--- program DoorRL_C (robot ABB IRB 1300-10/1.15) ---
  Smooth(1)
  Set speed (1000.0 mm/s)
  Set Ref.: DoorRL
  Set Tool: Generic Paint Sprayer
  Show Generic Paint Sprayer
  MoveJ 1 to (90.7, 0.32, 7.32) mm, rotated rx -9.04 ry 0.01 rz 91.21 deg; joints [83.599, -28.806, 2.512, -49.508, 32.312, -224.781, 2064.306, 3452.351, 803.193]
  MoveL 2 to (90.7, 0.32, 7.32) mm, rotated rx -9.04 ry 0.01 rz 91.21 deg; joints [83.599, -28.806, 2.512, -49.508, 32.312, -224.781, 2064.306, 3452.351, 803.193]
  MoveL 3 to (75, 0, 106.08) mm, rotated rx -9.04 ry 0.01 rz 91.21 deg; joints [85.387, -19.776, -1.909, -57.854, 30.896, -215.842, 2064.306, 3452.351, 803.193]
  MoveL 4 to (75, 0, 106.08) mm, rotated rx -9.04 ry 0.01 rz 91.21 deg; joints [85.387, -19.776, -1.909, -57.854, 30.896, -215.842, 2064.306, 3452.351, 803.193]
  Set speed (200.0 mm/s)
  MoveL 5 to (75, 100, 106.62) mm, rotated rx -8.72 ry -0.14 rz 91.23 deg; joints [102.46, -18.99, -2.4, -72.728, 45.516, -205.072, 2064.306, 3452.351, 803.193]
  MoveL 6 to (75, 200, 107.42) mm, rotated rx -8.48 ry -0.48 rz 91.28 deg; joints [117.629, -15.548, -4.305, -81.612, 59.424, -199.395, 2064.306, 3452.351, 803.193]
  MoveL 7 to (75, 300, 108.62) mm, rotated rx -8.1 ry -0.62 rz 91.29 deg; joints [129.26, -10.149, -8.101, -86.402, 70.427, -196.705, 2064.306, 3452.351, 803.193]
  MoveL 8 to (75, 400, 110.17) mm, rotated rx -8.3 ry -0.88 rz 91.34 deg; joints [137.912, -3.315, -13.206, -89.791, 78.836, -194.463, 2064.306, 3452.351, 803.193]
  MoveL 9 to (75, 500, 112.34) mm, rotated rx -7.79 ry -1.35 rz 91.39 deg; joints [144.305, 5.186, -22.224, -91.259, 85.516, -195.347, 2064.306, 3452.351, 803.193]
  MoveL 10 to (75, 600, 114.4) mm, rotated rx -6.61 ry -0.07 rz 91.2 deg; joints [148.976, 13.47, -33.602, -91.242, 88.944, -199.214, 2064.306, 3452.351, 803.193]
  Set speed (1000.0 mm/s)
  MoveL 11 to (75, 600, 114.4) mm, rotated rx -6.61 ry -0.07 rz 91.2 deg; joints [148.976, 13.47, -33.602, -91.242, 88.944, -199.214, 2064.306, 3452.351, 803.193]
  MoveL 12 to (86.51, 600.37, 15.07) mm, rotated rx -6.61 ry -0.07 rz 91.2 deg; joints [156.899, 8.317, -26.551, -93.775, 96.503, -197.647, 2064.306, 3452.351, 803.193]
  Set speed (1000.0 mm/s)
  MoveL 13 to (152.01, 598.2, 20.45) mm, rotated rx -1.13 ry 1.05 rz 91.14 deg; joints [156.743, 6.079, -21.228, -88.467, 96.739, -196.702, 2064.306, 3452.351, 803.193]
  MoveL 14 to (150, 600, 120.41) mm, rotated rx -1.13 ry 1.05 rz 91.14 deg; joints [148.769, 10.819, -26.045, -86.396, 89.056, -197.123, 2064.306, 3452.351, 803.193]
  MoveL 15 to (150, 600, 120.41) mm, rotated rx -1.13 ry 1.05 rz 91.14 deg; joints [148.769, 10.819, -26.045, -86.396, 89.056, -197.123, 2064.306, 3452.351, 803.193]
  Set speed (200.0 mm/s)
  MoveL 16 to (150, 500, 121.61) mm, rotated rx -2.1 ry 0.62 rz 91.14 deg; joints [143.656, 2.312, -15.23, -86.198, 84.142, -194.609, 2064.306, 3452.351, 803.193]
  MoveL 17 to (150, 400, 121.47) mm, rotated rx -4.4 ry -0.1 rz 91.19 deg; joints [137.209, -5.289, -5.416, -87.296, 77.972, -191.254, 2064.306, 3452.351, 803.193]
  MoveL 18 to (150, 300, 120.53) mm, rotated rx -8.5 ry -0.52 rz 91.29 deg; joints [128.581, -12.398, 4.736, -90.48, 69.312, -185.121, 2064.306, 3452.351, 803.193]
  MoveL 19 to (150, 200, 119.49) mm, rotated rx -8.12 ry -0.38 rz 91.26 deg; joints [116.951, -17.771, 7.428, -86.802, 57.781, -188.768, 2064.306, 3452.351, 803.193]
  MoveL 20 to (150, 100, 118.81) mm, rotated rx -7.65 ry -0.05 rz 91.21 deg; joints [101.911, -21.13, 8.356, -79.735, 43.178, -194.732, 2064.306, 3452.351, 803.193]
  MoveL 21 to (150, 0, 118.53) mm, rotated rx -7.91 ry 0.3 rz 91.16 deg; joints [84.752, -21.907, 8.755, -69.015, 26.732, -202.933, 2064.306, 3452.351, 803.193]
  Set speed (1000.0 mm/s)
  MoveL 22 to (150, 0, 118.53) mm, rotated rx -7.91 ry 0.3 rz 91.16 deg; joints [84.752, -21.907, 8.755, -69.015, 26.732, -202.933, 2064.306, 3452.351, 803.193]
  MoveL 23 to (163.76, -0.24, 19.48) mm, rotated rx -7.91 ry 0.3 rz 91.16 deg; joints [82.61, -31.376, 12.865, -57.206, 27.32, -215.521, 2064.306, 3452.351, 803.193]
  Set speed (1000.0 mm/s)
  MoveL 24 to (223.66, 0.79, 20.64) mm, rotated rx 0.76 ry -0.47 rz 91.14 deg; joints [84.141, -30.772, 10.615, -47.345, 35.088, -229.019, 2064.306, 3452.351, 803.193]
  MoveL 25 to (225, 0, 120.63) mm, rotated rx 0.76 ry -0.47 rz 91.14 deg; joints [85.606, -21.929, 8.883, -57.612, 31.856, -217.231, 2064.306, 3452.351, 803.193]
  MoveL 26 to (225, 0, 120.63) mm, rotated rx 0.76 ry -0.47 rz 91.14 deg; joints [85.606, -21.929, 8.883, -57.612, 31.856, -217.231, 2064.306, 3452.351, 803.193]
  Set speed (200.0 mm/s)
  MoveL 27 to (225, 100, 121.28) mm, rotated rx 0.7 ry -0.35 rz 91.14 deg; joints [102.099, -21.314, 8.944, -70.725, 45.982, -205.135, 2064.306, 3452.351, 803.193]
  MoveL 28 to (225, 200, 122.15) mm, rotated rx 0.5 ry -0.52 rz 91.15 deg; joints [117.028, -17.979, 7.742, -78.485, 59.657, -197.425, 2064.306, 3452.351, 803.193]
  MoveL 29 to (225, 300, 123.05) mm, rotated rx 0.21 ry -0.42 rz 91.15 deg; joints [128.604, -12.816, 5.114, -82.577, 70.367, -192.361, 2064.306, 3452.351, 803.193]
  MoveL 30 to (225, 400, 123.5) mm, rotated rx -0.2 ry -0.26 rz 91.16 deg; joints [137.37, -6.35, 0.883, -84.796, 78.558, -188.773, 2064.306, 3452.351, 803.193]
  MoveL 31 to (225, 500, 123.04) mm, rotated rx -1.05 ry 0.5 rz 91.15 deg; joints [143.943, 0.436, -4.189, -86.301, 84.114, -186.009, 2064.306, 3452.351, 803.193]
  MoveL 32 to (225, 600, 122.08) mm, rotated rx -1.6 ry 0.73 rz 91.14 deg; joints [149.099, 8.52, -12.229, -87.11, 88.967, -185.37, 2064.306, 3452.351, 803.193]
  MoveL 33 to (225, 700, 120.88) mm, rotated rx 0.16 ry -3.32 rz 91.14 deg; joints [153.063, 22.747, -33.337, -87.148, 97.49, -192.931, 2064.306, 3452.351, 803.193]
  Set speed (1000.0 mm/s)
  MoveL 34 to (225, 700, 120.88) mm, rotated rx 0.16 ry -3.32 rz 91.14 deg; joints [153.063, 22.747, -33.337, -87.148, 97.49, -192.931, 2064.306, 3452.351, 803.193]
  MoveL 35 to (224.61, 705.78, 21.05) mm, rotated rx 0.16 ry -3.32 rz 91.14 deg; joints [160.083, 19.015, -28.957, -88.222, 104.365, -191.988, 2064.306, 3452.351, 803.193]
  Set speed (1000.0 mm/s)
  MoveL 36 to (305.54, 698.73, 24.64) mm, rotated rx -3.16 ry 0.79 rz 91.13 deg; joints [160.573, 12.44, -5.322, -87.261, 99.896, -173.342, 2064.306, 3452.351, 803.193]
  MoveL 37 to (300, 700, 124.48) mm, rotated rx -3.16 ry 0.79 rz 91.13 deg; joints [153.278, 16.534, -10.403, -88.244, 92.694, -174.618, 2064.306, 3452.351, 803.193]
  MoveL 38 to (300, 700, 124.48) mm, rotated rx -3.16 ry 0.79 rz 91.13 deg; joints [153.278, 16.534, -10.403, -88.244, 92.694, -174.618, 2064.306, 3452.351, 803.193]
  Set speed (200.0 mm/s)
  MoveL 39 to (300, 600, 125.06) mm, rotated rx -3.23 ry 0.19 rz 91.16 deg; joints [149.376, 8.214, 0.141, -88.693, 89.372, -172.462, 2064.306, 3452.351, 803.193]
  MoveL 40 to (300, 500, 125.16) mm, rotated rx -2.17 ry 0.14 rz 91.16 deg; joints [144.303, -0.143, 7.785, -88.428, 84.307, -173.89, 2064.306, 3452.351, 803.193]
  MoveL 41 to (300, 400, 124.72) mm, rotated rx -1.66 ry -0.34 rz 91.17 deg; joints [137.782, -7.551, 13.671, -88.464, 78.321, -175.937, 2064.306, 3452.351, 803.193]
  MoveL 42 to (300, 300, 123.67) mm, rotated rx -1.09 ry -0.54 rz 91.17 deg; joints [129.056, -14.44, 17.858, -87.824, 69.893, -179.463, 2064.306, 3452.351, 803.193]
  MoveL 43 to (300, 200, 122.54) mm, rotated rx -1.3 ry -0.63 rz 91.18 deg; joints [117.411, -20.166, 21.239, -87.099, 58.454, -182.429, 2064.306, 3452.351, 803.193]
  MoveL 44 to (300, 100, 121.57) mm, rotated rx -1.33 ry -0.43 rz 91.17 deg; joints [102.223, -23.973, 22.85, -84.399, 43.259, -186.653, 2064.306, 3452.351, 803.193]
  MoveL 45 to (300, 0, 120.78) mm, rotated rx -1.5 ry -0.32 rz 91.17 deg; joints [85.014, -24.825, 23.131, -79.981, 26.14, -191.455, 2064.306, 3452.351, 803.193]
  Set speed (1000.0 mm/s)
  MoveL 46 to (300, 0, 120.78) mm, rotated rx -1.5 ry -0.32 rz 91.17 deg; joints [85.014, -24.825, 23.131, -79.981, 26.14, -191.455, 2064.306, 3452.351, 803.193]
  MoveL 47 to (302.6, 0.61, 20.82) mm, rotated rx -1.5 ry -0.32 rz 91.17 deg; joints [83.173, -35.007, 25.553, -63.775, 26.819, -209.331, 2064.306, 3452.351, 803.193]
  Set speed (1000.0 mm/s)
  MoveL 48 to (382.47, 0.73, 24.79) mm, rotated rx -4.29 ry -0.33 rz 91.21 deg; joints [82.724, -37.124, 40.086, -95.64, 23.549, -173.926, 2064.306, 3452.351, 803.193]
  MoveL 49 to (375, 0, 124.51) mm, rotated rx -4.29 ry -0.33 rz 91.21 deg; joints [84.717, -25.281, 36.632, -111.575, 27.492, -156.03, 2064.306, 3452.351, 803.193]
  MoveL 50 to (375, 0, 124.51) mm, rotated rx -4.29 ry -0.33 rz 91.21 deg; joints [84.717, -25.281, 36.632, -111.575, 27.492, -156.03, 2064.306, 3452.351, 803.193]
  Set speed (200.0 mm/s)
  MoveL 51 to (375, 100, 125.3) mm, rotated rx -4.19 ry -0.39 rz 91.21 deg; joints [102.046, -24.392, 36.412, -101.899, 43.99, -163.49, 2064.306, 3452.351, 803.193]
  MoveL 52 to (375, 200, 126.3) mm, rotated rx -3.97 ry -0.6 rz 91.22 deg; joints [117.418, -20.181, 34.415, -97.776, 59.26, -164.282, 2064.306, 3452.351, 803.193]
  MoveL 53 to (375, 300, 127.56) mm, rotated rx -5.31 ry -0.62 rz 91.24 deg; joints [129.232, -13.59, 32.312, -96.985, 71.452, -159.822, 2064.306, 3452.351, 803.193]
  MoveL 54 to (375, 400, 128.83) mm, rotated rx -5.27 ry -0.59 rz 91.24 deg; joints [137.993, -6.109, 26.861, -94.307, 79.819, -158.606, 2064.306, 3452.351, 803.193]
  MoveL 55 to (375, 500, 129.91) mm, rotated rx -4.47 ry -0.21 rz 91.2 deg; joints [144.445, 1.382, 19.151, -91.452, 85.235, -159.606, 2064.306, 3452.351, 803.193]
  MoveL 56 to (375, 600, 130.48) mm, rotated rx -5.59 ry -0.1 rz 91.2 deg; joints [149.411, 9.838, 11.165, -90.644, 90.13, -158.616, 2064.306, 3452.351, 803.193]
  MoveL 57 to (375, 700, 130.64) mm, rotated rx -6.1 ry 0.33 rz 91.16 deg; joints [153.257, 18.109, 1.02, -89.952, 93.484, -160.267, 2064.306, 3452.351, 803.193]
  MoveL 58 to (375, 800, 129.84) mm, rotated rx -6.14 ry 1.82 rz 91 deg; joints [156.376, 25.705, -10.148, -89.777, 95.052, -163.863, 2064.306, 3452.351, 803.193]
  Set speed (1000.0 mm/s)
  MoveL 59 to (375, 800, 129.84) mm, rotated rx -6.14 ry 1.82 rz 91 deg; joints [156.376, 25.705, -10.148, -89.777, 95.052, -163.863, 2064.306, 3452.351, 803.193]
  MoveL 60 to (385.74, 797.03, 30.46) mm, rotated rx -6.14 ry 1.82 rz 91 deg; joints [163.022, 22.035, -4.129, -87.501, 101.36, -161.341, 2064.306, 3452.351, 803.193]
  Set speed (1000.0 mm/s)
  MoveL 61 to (473.75, 798.92, 46.41) mm, rotated rx -13.73 ry 0.89 rz 91.03 deg; joints [161.964, 28.907, 7.054, -89.444, 104.008, -140.367, 2064.306, 3452.351, 803.193]
  MoveL 62 to (450, 800, 143.54) mm, rotated rx -13.73 ry 0.89 rz 91.03 deg; joints [155.503, 31.395, 0.291, -93.866, 98.516, -144.558, 2064.306, 3452.351, 803.193]
  MoveL 63 to (450, 800, 143.54) mm, rotated rx -13.73 ry 0.89 rz 91.03 deg; joints [155.503, 31.395, 0.291, -93.866, 98.516, -144.558, 2064.306, 3452.351, 803.193]
  Set speed (200.0 mm/s)
  MoveL 64 to (450, 700, 143.19) mm, rotated rx -13.87 ry 0.24 rz 91.18 deg; joints [152.373, 24.011, 12.763, -94.602, 96.91, -139.132, 2064.306, 3452.351, 803.193]
  MoveL 65 to (450, 600, 141.71) mm, rotated rx -14.05 ry -0.52 rz 91.38 deg; joints [148.554, 17.067, 23.436, -96.144, 94.968, -134.987, 2064.306, 3452.351, 803.193]
  MoveL 66 to (450, 500, 140.16) mm, rotated rx -13.37 ry -0.76 rz 91.42 deg; joints [143.712, 9.342, 32.755, -98.644, 91.321, -133.254, 2064.306, 3452.351, 803.193]
  MoveL 67 to (450, 400, 138.58) mm, rotated rx -12.7 ry -0.52 rz 91.35 deg; joints [137.185, 1.179, 40.884, -102.834, 85.962, -132.737, 2064.306, 3452.351, 803.193]
  MoveL 68 to (450, 300, 137.1) mm, rotated rx -11.58 ry -0.68 rz 91.37 deg; joints [128.567, -6.84, 46.323, -107.585, 78.404, -134.195, 2064.306, 3452.351, 803.193]
  MoveL 69 to (450, 200, 135.73) mm, rotated rx -11.11 ry -0.72 rz 91.37 deg; joints [116.912, -13.706, 50.251, -114.63, 68.528, -133.929, 2064.306, 3452.351, 803.193]
  MoveL 70 to (450, 100, 134.52) mm, rotated rx -9.69 ry -0.28 rz 91.26 deg; joints [101.492, -19.511, 51.351, -123.947, 53.928, -132.478, 2064.306, 3452.351, 803.193]
  MoveL 71 to (450, 0, 133.84) mm, rotated rx -9.43 ry -0.15 rz 91.24 deg; joints [84.256, -20.688, 51.274, -141.098, 41.917, -120.478, 2064.306, 3452.351, 803.193]
  Set speed (1000.0 mm/s)
  MoveL 72 to (450, 0, 133.84) mm, rotated rx -9.43 ry -0.15 rz 91.24 deg; joints [84.256, -20.688, 51.274, -141.098, 41.917, -120.478, 2064.306, 3452.351, 803.193]
  MoveL 73 to (466.37, 0.62, 35.19) mm, rotated rx -9.43 ry -0.15 rz 91.24 deg; joints [82.039, -34.232, 56.958, -137.497, 34.657, -126.322, 2064.306, 3452.351, 803.193]
  Set speed (1000.0 mm/s)
  MoveL 74 to (555.05, -82.25, 116.77) mm, rotated rx 60.29 ry -13.07 rz -152.57 deg; joints [70.284, 61.29, -33.097, 77.942, 86.027, -269.551, 2564.306, 3828.918, 1060.29]
  MoveL 75 to (525, 0, 165.05) mm, rotated rx 37.44 ry 52.55 rz 154.03 deg; joints [24.866, 61.421, -22.556, 79.321, 94.582, -359.342, 1755.93, 3452.351, 1099.978]
  MoveL 76 to (525, 0, 165.05) mm, rotated rx 37.44 ry 52.55 rz 154.03 deg; joints [24.866, 61.421, -22.556, 79.321, 94.582, -359.342, 1755.93, 3452.351, 1099.978]
  Set speed (200.0 mm/s)
  MoveL 77 to (525, 100, 155.04) mm, rotated rx -9.84 ry 16.5 rz 149.85 deg; joints [40.939, 27.228, 59.96, 145.73, 75.776, -387.964, 1755.93, 3452.351, 1099.978]
  MoveL 78 to (525, 200, 156.11) mm, rotated rx 15.18 ry 12.68 rz -126.97 deg; joints [110.817, 44.311, 23.812, 178.664, 63.101, -311.328, 2564.306, 3828.918, 1099.979]
  MoveL 79 to (525, 300, 157.73) mm, rotated rx -8.79 ry -16.06 rz 32.63 deg; joints [133.225, 83.406, -21.75, 229.016, 112.204, -168.506, 2564.306, 3742.832, 1099.974]
  MoveL 80 to (525, 400, 159.79) mm, rotated rx -8.89 ry -16.44 rz 32.7 deg; joints [137.126, 86.051, -37.16, 228.381, 105.823, -180.156, 2564.306, 3742.832, 1060.252]
  MoveL 81 to (525, 500, 162.03) mm, rotated rx -9.11 ry -16.87 rz 32.78 deg; joints [140.443, 100.168, -72.983, 227.152, 93.486, -198.143, 2564.306, 3742.832, 1060.252]
  MoveL 82 to (525, 600, 164.37) mm, rotated rx -9.81 ry -18.17 rz 33.04 deg; joints [119.482, 84.102, -18.159, 219.568, 113.288, -160.148, 2064.306, 3834.482, 1099.978]
  MoveL 83 to (525, 700, 166.85) mm, rotated rx -10.72 ry -19.05 rz 33.23 deg; joints [124.134, 85.187, -28.709, 220.198, 108.523, -168.206, 2064.306, 3834.482, 1060.086]
  MoveL 84 to (525, 800, 169.19) mm, rotated rx -11.61 ry -20.92 rz 33.67 deg; joints [131.809, 86.524, -29.394, 225.322, 113.849, -170.732, 2064.306, 3735.345, 1060.086]
  MoveL 85 to (525, 900, 171.75) mm, rotated rx -12.62 ry -22.91 rz 34.2 deg; joints [135.296, 97.473, -57.469, 222.496, 105.147, -184.837, 2064.306, 3735.345, 1060.086]
  Set speed (1000.0 mm/s)
  MoveL 86 to (525, 900, 171.75) mm, rotated rx -12.62 ry -22.91 rz 34.2 deg; joints [135.296, 97.473, -57.469, 222.496, 105.147, -184.837, 2064.306, 3735.345, 1060.086]
  MoveL 87 to (568.69, 903.29, 81.86) mm, rotated rx -12.62 ry -22.91 rz 34.2 deg; joints [135.12, 104.561, -69.901, 221.579, 101.084, -188.404, 2064.306, 3836.185, 1060.086]
  Set speed (1000.0 mm/s)
  MoveL 88 to (674.57, 902.94, 144.38) mm, rotated rx -46.41 ry -15.12 rz 78.31 deg; joints [105.449, 76.927, -11.434, 224.156, 120.066, -102.909, 1454.359, 3827.063, 803.193]
  MoveL 89 to (600, 900, 210.95) mm, rotated rx -46.41 ry -15.12 rz 78.31 deg; joints [105.243, 71.137, -8.955, 222.754, 117.599, -105.433, 1454.359, 3760.201, 803.193]
  MoveL 90 to (600, 900, 210.95) mm, rotated rx -46.41 ry -15.12 rz 78.31 deg; joints [105.243, 71.137, -8.955, 222.754, 117.599, -105.433, 1454.359, 3760.201, 803.193]
  Set speed (200.0 mm/s)
  MoveL 91 to (600, 800, 210) mm, rotated rx 6.16 ry 2.87 rz 71.3 deg; joints [100.8, 46.533, 29.485, 219.508, 78.715, -121.802, 1454.359, 3760.201, 1056.724]
  MoveL 92 to (600, 700, 203.49) mm, rotated rx -43.73 ry -14.25 rz 77.35 deg; joints [92.704, 90.414, -14.669, 216.98, 122.816, -93.221, 1454.359, 3760.201, 1056.724]
  MoveL 93 to (600, 600, 200.56) mm, rotated rx -44.05 ry -14.06 rz 77.17 deg; joints [85.887, 90.364, -14.403, 211.003, 122.369, -91.43, 1454.359, 3760.201, 1056.724]
  MoveL 94 to (600, 500, 198.23) mm, rotated rx -43.4 ry -13.95 rz 77.05 deg; joints [79.336, 89.984, -14.885, 205.125, 120.303, -90.613, 1454.359, 3760.201, 1056.724]
  MoveL 95 to (600, 400, 196.18) mm, rotated rx -44.51 ry 0.19 rz 91.33 deg; joints [104.974, 82.58, -3.734, 227.238, 116.231, -77.118, 1920.961, 3772.068, 1056.724]
  MoveL 96 to (600, 300, 194.65) mm, rotated rx -43.34 ry 0.41 rz 91.12 deg; joints [98.134, 80.928, 1.713, 221.6, 117.257, -74.136, 1920.961, 3772.068, 1056.724]
  MoveL 97 to (600, 200, 193.74) mm, rotated rx -42.2 ry 0.55 rz 90.99 deg; joints [90.952, 79.687, 4.868, 214.872, 117.373, -72.904, 1920.961, 3772.068, 1056.724]
  MoveL 98 to (600, 100, 193.19) mm, rotated rx -40.28 ry 0.54 rz 91.01 deg; joints [83.708, 78.061, 6.898, 207.528, 115.777, -73.221, 1920.961, 3772.068, 1056.724]
  Set speed (1000.0 mm/s)
  MoveL 99 to (600, 100, 193.19) mm, rotated rx -40.28 ry 0.54 rz 91.01 deg; joints [83.708, 78.061, 6.898, 207.528, 115.777, -73.221, 1920.961, 3772.068, 1056.724]
  MoveL 100 to (664.66, 100.42, 116.91) mm, rotated rx -40.28 ry 0.54 rz 91.01 deg; joints [83.431, 83.386, 6.777, 208.563, 120.365, -70.437, 1920.961, 3823.518, 1056.724]
  Set speed (1000.0 mm/s)
  MoveL 101 to (748.8, 402.34, 190.34) mm, rotated rx -47.59 ry -0.13 rz 91.7 deg; joints [105.259, 99.236, -20.482, 228.709, 118.671, -75.099, 1920.961, 3768.591, 1056.724]
  MoveL 102 to (675, 400, 257.78) mm, rotated rx -47.59 ry -0.13 rz 91.7 deg; joints [103.965, 94.987, -25.674, 224.332, 111.906, -82.4, 1920.961, 3768.591, 1056.724]
  MoveL 103 to (675, 400, 257.78) mm, rotated rx -47.59 ry -0.13 rz 91.7 deg; joints [103.965, 94.987, -25.674, 224.332, 111.906, -82.4, 1920.961, 3768.591, 1056.724]
  Set speed (200.0 mm/s)
  MoveL 104 to (675, 500, 261.5) mm, rotated rx -47.59 ry -0.25 rz 91.84 deg; joints [109.884, 97.185, -33.463, 227.815, 109.711, -88.385, 1920.961, 3768.591, 1056.724]
  MoveL 105 to (675, 600, 265.72) mm, rotated rx -44.04 ry -14.72 rz 77.83 deg; joints [86.509, 101.363, -35.436, 209.841, 113.733, -96.969, 1454.359, 3755.143, 1056.724]
  MoveL 106 to (675, 700, 270.37) mm, rotated rx -41.7 ry -14.36 rz 77.4 deg; joints [92.877, 99.524, -31.623, 214.934, 114.764, -99.411, 1454.359, 3755.143, 1056.724]
  MoveL 107 to (675, 800, 275.52) mm, rotated rx -37.38 ry -13.59 rz 76.58 deg; joints [99.465, 96.499, -26.735, 220.282, 114.038, -102.592, 1454.359, 3755.143, 1056.724]
  MoveL 108 to (675, 900, 280.97) mm, rotated rx -37.72 ry -1.38 rz 92.5 deg; joints [104.161, 95.633, -32.168, 224.415, 99.282, -91.601, 1420.961, 3825.258, 1099.805]
  MoveL 109 to (675, 1000, 287.24) mm, rotated rx -31.01 ry -12.9 rz 75.77 deg; joints [112.266, 94.902, -31.121, 229.795, 108.116, -113.99, 1454.359, 3755.143, 1056.724]
  Set speed (1000.0 mm/s)
  MoveL 110 to (675, 1000, 287.24) mm, rotated rx -31.01 ry -12.9 rz 75.77 deg; joints [112.266, 94.902, -31.121, 229.795, 108.116, -113.99, 1454.359, 3755.143, 1056.724]
  MoveL 111 to (729.64, 1005.88, 203.7) mm, rotated rx -25.34 ry -22.43 rz 57.28 deg; joints [118.128, 111.273, -49.466, 227.376, 116.936, -137.304, 1564.306, 3749.389, 1099.805]

--- program DoorFL_C (robot ABB IRB 1300-10/1.15) ---
  Smooth(1)
  Set speed (1000.0 mm/s)
  Set Ref.: DoorFL
  Set Tool: Generic Paint Sprayer
  Show Generic Paint Sprayer
  MoveJ 1 to (71.29, 9.92, 20.7) mm, rotated rx 1.8 ry -5.81 rz 93.26 deg; joints [-42.65, -30.194, 5.671, 93.562, 99.411, 24.312, 2956.487, 3047.951, 891.281]
  MoveL 2 to (71.29, 9.92, 20.7) mm, rotated rx 1.8 ry -5.81 rz 93.26 deg; joints [-42.65, -30.194, 5.671, 93.562, 99.411, 24.312, 2956.487, 3047.951, 891.281]
  MoveL 3 to (75, 0, 120.14) mm, rotated rx 1.8 ry -5.81 rz 93.26 deg; joints [-42.65, -30.194, 5.671, 93.562, 99.411, 24.312, 2961.047, 2948.065, 889.846]
  MoveL 4 to (75, 0, 120.14) mm, rotated rx 1.8 ry -5.81 rz 93.26 deg; joints [-42.65, -30.194, 5.671, 93.562, 99.411, 24.312, 2961.047, 2948.065, 889.846]
  Set speed (200.0 mm/s)
  MoveL 5 to (75, 100, 126.97) mm, rotated rx -3.91 ry -2.93 rz 93.33 deg; joints [-42.529, -30.194, 9.554, 98.562, 100.324, 24.312, 2875.19, 2948.065, 860.651]
  MoveL 6 to (75, 200, 131.93) mm, rotated rx -5.64 ry -2.28 rz 93.25 deg; joints [-42.357, -30.194, 10.675, 99.97, 100.324, 24.312, 2777.783, 2947.743, 847.202]
  MoveL 7 to (75, 300, 136.32) mm, rotated rx -5.77 ry -2.17 rz 93.24 deg; joints [-42.357, -30.194, 10.767, 100.106, 100.386, 24.312, 2678.543, 2948.883, 840.768]
  MoveL 8 to (75, 400, 140.74) mm, rotated rx -5.66 ry -2.28 rz 93.25 deg; joints [-42.432, -30.263, 10.767, 100.006, 100.386, 24.312, 2578.494, 2949.946, 835.842]
  MoveL 9 to (75, 500, 145.36) mm, rotated rx -5.57 ry -2.46 rz 93.27 deg; joints [-42.582, -30.306, 10.767, 99.924, 100.386, 24.312, 2477.83, 2950.073, 830.733]
  MoveL 10 to (75, 600, 150.28) mm, rotated rx -5.46 ry -2.6 rz 93.29 deg; joints [-42.694, -30.37, 10.767, 99.824, 100.386, 24.312, 2377.497, 2950.334, 825.812]
  MoveL 11 to (75, 700, 155.46) mm, rotated rx -5.27 ry -2.81 rz 93.31 deg; joints [-42.844, -30.483, 10.767, 99.658, 100.386, 24.312, 2277.163, 2950.452, 821.515]
  MoveL 12 to (75, 800, 160.96) mm, rotated rx -5.04 ry -2.89 rz 93.32 deg; joints [-42.859, -30.634, 10.767, 99.472, 100.386, 24.312, 2177.86, 2951.505, 817.446]
  MoveL 13 to (75, 900, 166.78) mm, rotated rx -4.84 ry -3.09 rz 93.34 deg; joints [-43.002, -30.755, 10.767, 99.302, 100.386, 24.312, 2077.572, 2951.075, 813.21]
  MoveL 14 to (75, 1000, 172.94) mm, rotated rx -4.96 ry -3.25 rz 93.35 deg; joints [-43.002, -30.755, 10.829, 99.315, 100.205, 24.312, 1976.003, 2949.512, 806.878]
  Set speed (1000.0 mm/s)
  MoveL 15 to (75, 1000, 172.94) mm, rotated rx -4.96 ry -3.25 rz 93.35 deg; joints [-43.002, -30.755, 10.829, 99.315, 100.205, 24.312, 1976.003, 2949.512, 806.878]
  MoveL 16 to (83.3, 1006.15, 73.47) mm, rotated rx -4.96 ry -3.25 rz 93.35 deg; joints [-43.002, -30.755, 10.829, 99.315, 100.205, 24.312, 1975.903, 3048.977, 796.55]
  Set speed (1000.0 mm/s)
  MoveL 17 to (138.12, 1006, 73.54) mm, rotated rx 6.61 ry -3.85 rz 93.27 deg; joints [-43.002, -30.755, 4.046, 91.135, 103.088, 23.437, 1991.83, 3062.191, 796.55]
  MoveL 18 to (150, 1000, 172.65) mm, rotated rx 6.61 ry -3.85 rz 93.27 deg; joints [-43.002, -30.755, 4.046, 91.135, 103.088, 23.437, 1992.978, 2962.682, 786.723]
  MoveL 19 to (150, 1000, 172.65) mm, rotated rx 6.61 ry -3.85 rz 93.27 deg; joints [-43.002, -30.755, 4.046, 91.135, 103.088, 23.437, 1992.978, 2962.682, 786.723]
  Set speed (200.0 mm/s)
  MoveL 20 to (150, 900, 166.71) mm, rotated rx 6.33 ry -3.62 rz 93.3 deg; joints [-42.862, -30.547, 4.046, 91.347, 103.088, 23.437, 2092.73, 2962.933, 790.506]
  MoveL 21 to (150, 800, 161.05) mm, rotated rx 6.69 ry -3.59 rz 93.3 deg; joints [-42.862, -30.547, 3.806, 91.122, 103.228, 23.437, 2193.623, 2963.568, 797.896]
  MoveL 22 to (150, 700, 155.46) mm, rotated rx 6.83 ry -3.53 rz 93.31 deg; joints [-42.862, -30.547, 3.72, 91.057, 103.332, 23.437, 2294.406, 2964.045, 804.378]
  MoveL 23 to (150, 600, 150.01) mm, rotated rx 6.58 ry -3.37 rz 93.32 deg; joints [-42.79, -30.371, 3.72, 91.243, 103.332, 23.437, 2393.918, 2963.55, 808.425]
  MoveL 24 to (150, 500, 144.8) mm, rotated rx 6.55 ry -3.36 rz 93.33 deg; joints [-42.79, -30.346, 3.72, 91.271, 103.33, 23.437, 2493.74, 2963.138, 813.994]
  MoveL 25 to (150, 400, 139.67) mm, rotated rx 6.34 ry -3.25 rz 93.34 deg; joints [-42.746, -30.198, 3.72, 91.432, 103.33, 23.437, 2593.211, 2962.281, 818.301]
  MoveL 26 to (150, 300, 134.64) mm, rotated rx 6.25 ry -3.4 rz 93.32 deg; joints [-42.746, -30.169, 3.72, 91.432, 103.153, 23.453, 2691.526, 2961.021, 823.366]
  MoveL 27 to (150, 200, 129.17) mm, rotated rx 6.05 ry -3.86 rz 93.27 deg; joints [-42.746, -30.169, 3.72, 91.417, 102.663, 23.557, 2787.597, 2959.352, 827.234]
  MoveL 28 to (150, 100, 122.33) mm, rotated rx 6.08 ry -4.56 rz 93.2 deg; joints [-42.746, -30.169, 3.641, 91.123, 102.022, 23.557, 2881.855, 2958.013, 832.522]
  MoveL 29 to (150, 0, 113.92) mm, rotated rx 4.76 ry -5.25 rz 93.17 deg; joints [-42.746, -30.169, 4.475, 91.726, 100.959, 23.557, 2973.758, 2956.707, 832.182]
  Set speed (1000.0 mm/s)
  MoveL 30 to (150, 0, 113.92) mm, rotated rx 4.76 ry -5.25 rz 93.17 deg; joints [-42.746, -30.169, 4.475, 91.726, 100.959, 23.557, 2973.758, 2956.707, 832.182]
  MoveL 31 to (141.22, 8.65, 14.68) mm, rotated rx 4.76 ry -5.25 rz 93.17 deg; joints [-42.746, -30.169, 4.475, 91.726, 100.959, 23.557, 2970.16, 3056.425, 838.758]
  Set speed (1000.0 mm/s)
  MoveL 32 to (218.38, 6.67, 7.88) mm, rotated rx 3.57 ry -4.04 rz 93.29 deg; joints [-41.886, -28.581, 4.475, 92.48, 100.959, 22.798, 2970.26, 3056.429, 754.428]
  MoveL 33 to (225, 0, 107.44) mm, rotated rx 3.57 ry -4.04 rz 93.29 deg; joints [-41.886, -28.581, 4.475, 92.48, 100.959, 22.798, 2971.739, 2956.542, 749.901]
  MoveL 34 to (225, 0, 107.44) mm, rotated rx 3.57 ry -4.04 rz 93.29 deg; joints [-41.886, -28.581, 4.475, 92.48, 100.959, 22.798, 2971.739, 2956.542, 749.901]
  Set speed (200.0 mm/s)
  MoveL 35 to (225, 100, 114.85) mm, rotated rx 4.65 ry -4.66 rz 93.23 deg; joints [-42.149, -29.254, 4.399, 91.621, 100.959, 22.798, 2873.574, 2956.542, 751.585]
  MoveL 36 to (225, 200, 121.21) mm, rotated rx 5.64 ry -3.55 rz 93.31 deg; joints [-42.149, -29.398, 3.974, 91.38, 102.303, 22.797, 2785.609, 2961.897, 751.585]
  MoveL 37 to (225, 300, 126.42) mm, rotated rx 5.52 ry -3.08 rz 93.36 deg; joints [-42.149, -29.398, 4.093, 91.637, 102.695, 22.797, 2689.308, 2963.788, 745.623]
  MoveL 38 to (225, 400, 131.18) mm, rotated rx 5.51 ry -3.04 rz 93.36 deg; joints [-42.149, -29.398, 4.103, 91.66, 102.731, 22.797, 2589.703, 2964.649, 739.767]
  MoveL 39 to (225, 500, 136.13) mm, rotated rx 5.58 ry -3.21 rz 93.34 deg; joints [-42.292, -29.461, 4.103, 91.606, 102.731, 22.798, 2489.295, 2964.561, 734.446]
  MoveL 40 to (225, 600, 141.25) mm, rotated rx 5.36 ry -3.25 rz 93.34 deg; joints [-42.292, -29.461, 4.25, 91.74, 102.614, 22.798, 2388.505, 2964.499, 727.583]
  MoveL 41 to (225, 700, 146.61) mm, rotated rx 5.44 ry -3.42 rz 93.32 deg; joints [-42.437, -29.525, 4.25, 91.683, 102.614, 22.798, 2288.064, 2963.987, 722.289]
  MoveL 42 to (225, 800, 152.19) mm, rotated rx 5.47 ry -3.55 rz 93.31 deg; joints [-42.553, -29.55, 4.25, 91.668, 102.614, 22.798, 2187.583, 2963.245, 716.614]
  MoveL 43 to (225, 900, 158) mm, rotated rx 5.36 ry -3.68 rz 93.3 deg; joints [-42.553, -29.55, 4.31, 91.69, 102.458, 22.798, 2086.278, 2962.296, 710.213]
  MoveL 44 to (225, 1000, 164.01) mm, rotated rx 5.47 ry -3.81 rz 93.29 deg; joints [-42.651, -29.633, 4.31, 91.607, 102.458, 22.798, 1986.16, 2961.565, 705.174]
  Set speed (1000.0 mm/s)
  MoveL 45 to (225, 1000, 164.01) mm, rotated rx 5.47 ry -3.81 rz 93.29 deg; joints [-42.651, -29.633, 4.31, 91.607, 102.458, 22.798, 1986.16, 2961.565, 705.174]
  MoveL 46 to (215.1, 1006.06, 64.69) mm, rotated rx 5.47 ry -3.81 rz 93.29 deg; joints [-42.651, -29.633, 4.31, 91.607, 102.458, 22.798, 1985.083, 3061.251, 713.019]
  Set speed (1000.0 mm/s)
  MoveL 47 to (294.37, 1006.17, 58.43) mm, rotated rx 3.02 ry -3.72 rz 93.32 deg; joints [-42.651, -29.454, 5.768, 93.281, 101.791, 22.798, 1985.083, 3062.29, 622.549]
  MoveL 48 to (300, 1000, 158.08) mm, rotated rx 3.02 ry -3.72 rz 93.32 deg; joints [-42.651, -29.454, 5.768, 93.281, 101.791, 22.798, 1986.004, 2962.358, 618.975]
  MoveL 49 to (300, 1000, 158.08) mm, rotated rx 3.02 ry -3.72 rz 93.32 deg; joints [-42.651, -29.454, 5.768, 93.281, 101.791, 22.798, 1986.004, 2962.358, 618.975]
  Set speed (200.0 mm/s)
  MoveL 50 to (300, 900, 151.94) mm, rotated rx 3.06 ry -3.64 rz 93.32 deg; joints [-42.646, -29.454, 5.746, 93.281, 101.873, 22.798, 2086.746, 2963.398, 625.029]
  MoveL 51 to (300, 800, 146.05) mm, rotated rx 3.14 ry -3.47 rz 93.33 deg; joints [-42.614, -29.454, 5.705, 93.281, 102.034, 22.797, 2188.302, 2964.697, 631.316]
  MoveL 52 to (300, 700, 140.44) mm, rotated rx 3.09 ry -3.31 rz 93.34 deg; joints [-42.469, -29.416, 5.705, 93.317, 102.034, 22.797, 2288.9, 2965.619, 636.801]
  MoveL 53 to (300, 600, 135.08) mm, rotated rx 3.06 ry -3.16 rz 93.35 deg; joints [-42.331, -29.393, 5.705, 93.336, 102.034, 22.797, 2389.526, 2966.32, 642.458]
  MoveL 54 to (300, 500, 129.95) mm, rotated rx 3.38 ry -3.11 rz 93.35 deg; joints [-42.33, -29.393, 5.498, 93.137, 102.175, 22.797, 2490.464, 2966.57, 649.722]
  MoveL 55 to (300, 400, 125.04) mm, rotated rx 3.59 ry -2.96 rz 93.36 deg; joints [-42.33, -29.393, 5.374, 93.055, 102.382, 22.797, 2592.092, 2966.844, 656.583]
  MoveL 56 to (300, 300, 120.32) mm, rotated rx 3.73 ry -2.91 rz 93.36 deg; joints [-42.238, -29.393, 5.28, 92.938, 102.382, 22.797, 2692.413, 2966.728, 663.053]
  MoveL 57 to (300, 200, 115.54) mm, rotated rx 2.72 ry -2.93 rz 93.36 deg; joints [-42.238, -29.102, 5.651, 93.618, 102.062, 22.797, 2788.523, 2962.966, 663.053]
  MoveL 58 to (300, 100, 109.76) mm, rotated rx 2.23 ry -4.12 rz 93.31 deg; joints [-42.238, -29.102, 5.651, 93.546, 100.793, 23.034, 2878.261, 2958.593, 664.498]
  MoveL 59 to (300, 0, 103.13) mm, rotated rx 1.82 ry -3.32 rz 93.34 deg; joints [-41.557, -28.818, 5.651, 93.866, 100.793, 23.034, 2980.655, 2962.9, 667.356]
  Set speed (1000.0 mm/s)
  MoveL 60 to (300, 0, 103.13) mm, rotated rx 1.82 ry -3.32 rz 93.34 deg; joints [-41.557, -28.818, 5.651, 93.866, 100.793, 23.034, 2980.655, 2962.9, 667.356]
  MoveL 61 to (296.5, 5.59, 3.35) mm, rotated rx 1.82 ry -3.32 rz 93.34 deg; joints [-41.557, -28.818, 5.651, 93.866, 100.793, 23.034, 2980.443, 3062.889, 668.834]
  Set speed (1000.0 mm/s)
  MoveL 62 to (376.58, 7.63, 2.13) mm, rotated rx -1.16 ry -4.32 rz 93.37 deg; joints [-41.557, -28.818, 7.489, 95.543, 99.023, 23.034, 2969.852, 3054.063, 575.476]
  MoveL 63 to (375, 0, 101.83) mm, rotated rx -1.16 ry -4.32 rz 93.37 deg; joints [-41.557, -28.818, 7.489, 95.543, 99.023, 23.034, 2971.805, 2954.151, 579.192]
  MoveL 64 to (375, 0, 101.83) mm, rotated rx -1.16 ry -4.32 rz 93.37 deg; joints [-41.557, -28.818, 7.489, 95.543, 99.023, 23.034, 2971.805, 2954.151, 579.192]
  Set speed (200.0 mm/s)
  MoveL 65 to (375, 100, 108.61) mm, rotated rx -1.56 ry -3.05 rz 93.34 deg; joints [-41.557, -28.818, 7.828, 96.312, 100.084, 23.034, 2881.73, 2957.046, 571.975]
  MoveL 66 to (375, 200, 113.89) mm, rotated rx -0.83 ry -2.73 rz 93.34 deg; joints [-41.557, -29.259, 7.828, 95.927, 100.585, 23.034, 2788.557, 2962.292, 571.594]
  MoveL 67 to (375, 300, 118.55) mm, rotated rx -1.03 ry -2.48 rz 93.33 deg; joints [-41.557, -29.259, 7.971, 96.16, 100.76, 23.034, 2690.4, 2963.686, 564.962]
  MoveL 68 to (375, 400, 123.13) mm, rotated rx -1.16 ry -2.66 rz 93.33 deg; joints [-41.557, -29.259, 8.041, 96.181, 100.555, 23.034, 2588.716, 2963.676, 558.469]
  MoveL 69 to (375, 500, 128.02) mm, rotated rx -1.34 ry -2.8 rz 93.34 deg; joints [-41.557, -29.259, 8.147, 96.255, 100.375, 23.034, 2487.297, 2963.424, 551.775]
  MoveL 70 to (375, 600, 133.18) mm, rotated rx -1.32 ry -2.99 rz 93.34 deg; joints [-41.739, -29.268, 8.147, 96.231, 100.375, 23.034, 2386.306, 2962.482, 546.142]
  MoveL 71 to (375, 700, 138.67) mm, rotated rx -1.29 ry -3.17 rz 93.34 deg; joints [-41.908, -29.283, 8.147, 96.201, 100.375, 23.034, 2285.414, 2961.353, 540.574]
  MoveL 72 to (375, 800, 144.43) mm, rotated rx -1.29 ry -3.3 rz 93.35 deg; joints [-42.039, -29.283, 8.153, 96.2, 100.375, 23.034, 2184.652, 2960.099, 534.778]
  MoveL 73 to (375, 900, 150.42) mm, rotated rx -1.35 ry -3.44 rz 93.35 deg; joints [-42.073, -29.283, 8.185, 96.2, 100.263, 23.034, 2083.478, 2958.84, 528.675]
  MoveL 74 to (375, 1000, 156.73) mm, rotated rx -1.55 ry -3.61 rz 93.36 deg; joints [-42.073, -29.283, 8.297, 96.269, 100.054, 23.034, 1981.723, 2957.006, 521.971]
  Set speed (1000.0 mm/s)
  MoveL 75 to (375, 1000, 156.73) mm, rotated rx -1.55 ry -3.61 rz 93.36 deg; joints [-42.073, -29.283, 8.297, 96.269, 100.054, 23.034, 1981.723, 2957.006, 521.971]
  MoveL 76 to (377.33, 1006.44, 56.97) mm, rotated rx -1.55 ry -3.61 rz 93.36 deg; joints [-42.073, -29.283, 8.297, 96.269, 100.054, 23.034, 1980.998, 3056.907, 517.58]
  Set speed (1000.0 mm/s)
  MoveL 77 to (468.92, 1006.72, 65.56) mm, rotated rx -11.12 ry -3.27 rz 93.36 deg; joints [-42.073, -29.284, 14.364, 103.155, 98.148, 23.034, 1975.183, 3025.414, 386.24]
  MoveL 78 to (450, 1000, 163.52) mm, rotated rx -11.12 ry -3.27 rz 93.36 deg; joints [-42.073, -29.284, 14.364, 103.155, 98.148, 23.034, 1975.321, 2927.631, 407.18]
  MoveL 79 to (450, 1000, 163.52) mm, rotated rx -11.12 ry -3.27 rz 93.36 deg; joints [-42.073, -29.284, 14.364, 103.155, 98.148, 23.034, 1975.321, 2927.631, 407.18]
  Set speed (200.0 mm/s)
  MoveL 80 to (450, 900, 156.95) mm, rotated rx -11.46 ry -3.12 rz 93.33 deg; joints [-41.991, -29.09, 14.364, 103.447, 98.148, 23.047, 2074.867, 2927.539, 410.366]
  MoveL 81 to (450, 800, 150.71) mm, rotated rx -11.88 ry -3.01 rz 93.31 deg; joints [-41.974, -28.826, 14.365, 103.785, 98.148, 23.047, 2173.519, 2925.972, 413.139]
  MoveL 82 to (450, 700, 144.66) mm, rotated rx -11.57 ry -2.7 rz 93.24 deg; joints [-41.974, -28.826, 14.194, 103.69, 98.505, 23.047, 2276.613, 2928.636, 420.053]
  MoveL 83 to (450, 600, 138.88) mm, rotated rx -10.26 ry -2.59 rz 93.24 deg; joints [-41.974, -28.826, 13.385, 102.792, 98.865, 23.047, 2379.103, 2933.078, 431.205]
  MoveL 84 to (450, 500, 133.53) mm, rotated rx -9.76 ry -2.56 rz 93.24 deg; joints [-41.974, -28.826, 13.071, 102.441, 98.995, 23.047, 2479.938, 2934.45, 439.13]
  MoveL 85 to (450, 400, 128.54) mm, rotated rx -9.61 ry -2.33 rz 93.2 deg; joints [-41.974, -28.826, 12.994, 102.427, 99.245, 23.047, 2582.083, 2935.231, 445.518]
  MoveL 86 to (450, 300, 123.82) mm, rotated rx -9.27 ry -2.27 rz 93.19 deg; joints [-41.974, -28.826, 12.783, 102.204, 99.373, 23.047, 2682.963, 2935.621, 452.792]
  MoveL 87 to (450, 200, 119.27) mm, rotated rx -9.13 ry -2.15 rz 93.18 deg; joints [-41.939, -28.826, 12.702, 102.147, 99.479, 23.047, 2783.994, 2935.621, 459.12]
  MoveL 88 to (450, 100, 114.42) mm, rotated rx -9.14 ry -2.59 rz 93.25 deg; joints [-41.939, -28.826, 12.674, 101.977, 99.064, 23.047, 2880.157, 2933.37, 465.059]
  MoveL 89 to (450, 0, 108.29) mm, rotated rx -9.36 ry -3.46 rz 93.39 deg; joints [-41.939, -28.826, 12.674, 101.799, 98.182, 23.125, 2972.591, 2930.297, 469.702]
  Set speed (1000.0 mm/s)
  MoveL 90 to (450, 0, 108.29) mm, rotated rx -9.36 ry -3.46 rz 93.39 deg; joints [-41.939, -28.826, 12.674, 101.799, 98.182, 23.125, 2972.591, 2930.297, 469.702]
  MoveL 91 to (465.88, 6.9, 9.8) mm, rotated rx -9.36 ry -3.46 rz 93.39 deg; joints [-41.939, -28.826, 12.674, 101.799, 98.182, 23.125, 2972.131, 3028.676, 451.778]
  Set speed (1000.0 mm/s)
  MoveL 92 to (572.67, 5.62, 33.94) mm, rotated rx -28.61 ry -2.16 rz 92.78 deg; joints [-41.939, -28.826, 24.837, 116.458, 96.895, 23.125, 2972.835, 2934.91, 275.292]
  MoveL 93 to (525, 0, 121.66) mm, rotated rx -28.61 ry -2.16 rz 92.78 deg; joints [-41.939, -28.826, 24.837, 116.458, 96.895, 23.125, 2970.772, 2847.987, 324.691]
  MoveL 94 to (525, 0, 121.66) mm, rotated rx -28.61 ry -2.16 rz 92.78 deg; joints [-41.939, -28.826, 24.837, 116.458, 96.895, 23.125, 2970.772, 2847.987, 324.691]
  Set speed (200.0 mm/s)
  MoveL 95 to (525, 100, 127.42) mm, rotated rx -7.04 ry -2.16 rz 93.22 deg; joints [-41.939, -28.826, 11.314, 100.665, 99.91, 23.125, 2890.372, 2925.932, 398.679]
  MoveL 96 to (525, 200, 131.94) mm, rotated rx -7.19 ry -2.22 rz 93.22 deg; joints [-42.033, -28.826, 11.416, 100.77, 99.908, 23.125, 2789.95, 2925.932, 392.331]
  MoveL 97 to (525, 300, 136.72) mm, rotated rx -8.29 ry -2.32 rz 93.22 deg; joints [-42.033, -28.826, 12.099, 101.513, 99.571, 23.125, 2687.705, 2923.516, 381.82]
  MoveL 98 to (525, 400, 141.76) mm, rotated rx -8.28 ry -2.43 rz 93.23 deg; joints [-42.137, -28.826, 12.109, 101.496, 99.57, 23.125, 2587.101, 2923.162, 376.158]
  MoveL 99 to (525, 500, 147.08) mm, rotated rx -8.24 ry -2.59 rz 93.26 deg; joints [-42.277, -28.839, 12.109, 101.442, 99.57, 23.125, 2486.321, 2922.399, 370.794]
  MoveL 100 to (525, 600, 152.91) mm, rotated rx 1.02 ry -3.42 rz 93.34 deg; joints [-42.277, -28.839, 6.141, 94.673, 101.128, 23.125, 2393.092, 2937.836, 404.369]
  MoveL 101 to (525, 700, 158.77) mm, rotated rx 1.05 ry -3.55 rz 93.34 deg; joints [-42.401, -28.86, 6.141, 94.648, 101.128, 23.125, 2292.496, 2936.69, 398.77]
  MoveL 102 to (525, 800, 164.86) mm, rotated rx 1.06 ry -3.63 rz 93.34 deg; joints [-42.477, -28.868, 6.141, 94.64, 101.128, 23.125, 2192.092, 2935.573, 393.025]
  MoveL 103 to (525, 900, 190.96) mm, rotated rx -1.81 ry -6.29 rz 93.44 deg; joints [-42.477, -28.868, 7.831, 95.569, 97.876, 23.125, 2064.179, 2899.315, 374.751]
  MoveL 104 to (525, 1000, 192.88) mm, rotated rx 3.5 ry 6.47 rz 93.93 deg; joints [-39.349, -28.868, 5.376, 95.569, 108.362, 23.125, 2074.244, 2962.879, 398.818]
  Set speed (1000.0 mm/s)
  MoveL 105 to (525, 1000, 192.88) mm, rotated rx 3.5 ry 6.47 rz 93.93 deg; joints [-39.349, -28.868, 5.376, 95.569, 108.362, 23.125, 2074.244, 2962.879, 398.818]
  MoveL 106 to (519.68, 988.35, 93.7) mm, rotated rx 3.5 ry 6.47 rz 93.93 deg; joints [-39.349, -28.868, 5.376, 95.569, 108.362, 23.125, 2091.074, 3061.358, 403.138]
  Set speed (1000.0 mm/s)
  MoveL 107 to (644.61, 1106.62, 141.81) mm, rotated rx -26.68 ry -2.69 rz 93.09 deg; joints [-52.744, -28.868, 28.66, 115.292, 108.357, 23.125, 1906.947, 2851.823, 184.092]
  MoveL 108 to (600, 1100, 231.06) mm, rotated rx -26.68 ry -2.69 rz 93.09 deg; joints [-52.744, -28.868, 28.66, 115.292, 108.357, 23.125, 1905.965, 2763.259, 230.518]
  MoveL 109 to (600, 1100, 231.06) mm, rotated rx -26.68 ry -2.69 rz 93.09 deg; joints [-52.744, -28.868, 28.66, 115.292, 108.357, 23.125, 1905.965, 2763.259, 230.518]
  Set speed (200.0 mm/s)
  MoveL 110 to (600, 1000, 223.62) mm, rotated rx -26.23 ry -2.68 rz 93.09 deg; joints [-52.733, -28.868, 28.302, 115.027, 108.361, 23.125, 2006.303, 2767.296, 237.066]
  MoveL 111 to (600, 900, 216.34) mm, rotated rx -26.2 ry -2.66 rz 93.08 deg; joints [-52.713, -28.868, 28.27, 115.016, 108.364, 23.125, 2106.535, 2769.394, 242.844]
  MoveL 112 to (600, 800, 209.28) mm, rotated rx -26.11 ry -2.47 rz 92.99 deg; joints [-52.529, -28.868, 28.143, 115.038, 108.365, 23.125, 2207.698, 2772.69, 248.023]
  MoveL 113 to (600, 700, 202.52) mm, rotated rx -25.61 ry -2.28 rz 92.9 deg; joints [-52.424, -28.868, 27.731, 114.813, 108.461, 23.125, 2309.355, 2777.238, 254.262]
  MoveL 114 to (600, 600, 196.18) mm, rotated rx -25.63 ry -2.11 rz 92.82 deg; joints [-52.264, -28.868, 27.699, 114.89, 108.461, 23.125, 2410.311, 2779.151, 259.37]
  MoveL 115 to (600, 500, 190.17) mm, rotated rx -26.01 ry -1.98 rz 92.75 deg; joints [-52.181, -28.709, 27.699, 115.218, 108.461, 23.245, 2510.371, 2777.748, 262.372]
  MoveL 116 to (600, 400, 184.44) mm, rotated rx -25.85 ry -1.86 rz 92.7 deg; joints [-52.095, -28.709, 27.557, 115.172, 108.498, 23.245, 2611.239, 2779.416, 268.114]
  MoveL 117 to (600, 300, 178.95) mm, rotated rx -23.63 ry -1.89 rz 92.77 deg; joints [-52.098, -28.709, 25.816, 113.784, 108.498, 23.245, 2711.759, 2788.958, 278.614]
  MoveL 118 to (600, 200, 173.63) mm, rotated rx -24.1 ry -1.79 rz 92.71 deg; joints [-52.097, -28.565, 25.816, 114.19, 108.498, 23.473, 2811.855, 2786.341, 280.918]
  MoveL 119 to (600, 100, 168.46) mm, rotated rx -25.05 ry -1.61 rz 92.6 deg; joints [-51.943, -27.896, 25.847, 114.847, 108.498, 23.473, 2908.86, 2778.394, 280.918]
  Set speed (1000.0 mm/s)
  MoveL 120 to (600, 100, 168.46) mm, rotated rx -25.05 ry -1.61 rz 92.6 deg; joints [-51.943, -27.896, 25.847, 114.847, 108.498, 23.473, 2908.86, 2778.394, 280.918]
  MoveL 121 to (642.19, 104.47, 77.9) mm, rotated rx -25.05 ry -1.61 rz 92.6 deg; joints [-51.943, -27.896, 25.847, 114.847, 108.498, 23.473, 2911.909, 2868.19, 237.017]

--- program DoorFR_C (robot ABB IRB 1300-10/1.15) ---
  Smooth(1)
  Set speed (1000.0 mm/s)
  Set Ref.: DoorFR
  Set Tool: Generic Paint Sprayer
  Show Generic Paint Sprayer
  MoveJ 1 to (-60.57, 1000.41, 143.85) mm, rotated rx 37.26 ry 1.12 rz 88.14 deg; joints [-120.367, 75.627, 1.596, -58.254, -113.465, 264.253, 2575.49, -300.668, 966.829]
  MoveL 2 to (-60.57, 1000.41, 143.85) mm, rotated rx 37.26 ry 1.12 rz 88.14 deg; joints [-120.367, 75.627, 1.596, -58.254, -113.465, 264.253, 2575.49, -300.668, 966.829]
  MoveL 3 to (0, 1000, 223.42) mm, rotated rx 37.26 ry 1.12 rz 88.14 deg; joints [-117.877, 73.425, -7.843, -52.577, -106.185, 273.954, 2575.49, -300.668, 966.829]
  MoveL 4 to (0, 1000, 223.42) mm, rotated rx 37.26 ry 1.12 rz 88.14 deg; joints [-117.877, 73.425, -7.843, -52.577, -106.185, 273.954, 2575.49, -300.668, 966.829]
  Set speed (200.0 mm/s)
  MoveL 5 to (0, 900, 222.5) mm, rotated rx 36.91 ry 0.93 rz 87.99 deg; joints [-112.228, 70.756, 0.07, -49.222, -107.556, 268.421, 2575.49, -300.668, 966.829]
  MoveL 6 to (0, 800, 221.68) mm, rotated rx 36.44 ry 0.96 rz 88 deg; joints [-105.926, 68.677, 6.264, -44.528, -108.61, 264.178, 2575.49, -300.668, 966.829]
  MoveL 7 to (0, 700, 221.06) mm, rotated rx 36.2 ry 1.08 rz 88.09 deg; joints [-99.072, 67.329, 10.29, -38.711, -109.338, 261.194, 2575.49, -300.668, 966.829]
  MoveL 8 to (0, 600, 220.88) mm, rotated rx 35.4 ry 1.2 rz 88.15 deg; joints [-91.927, 65.947, 12.846, -32.103, -108.773, 259.693, 2575.49, -300.668, 966.829]
  MoveL 9 to (0, 500, 220.39) mm, rotated rx 33.84 ry 0.88 rz 87.91 deg; joints [-84.962, 64.23, 14.029, -25.728, -106.23, 259.403, 2575.49, -300.668, 966.829]
  MoveL 10 to (0, 400, 220.95) mm, rotated rx 35.47 ry 1.81 rz 88.59 deg; joints [-77.269, 65.827, 10.349, -17.566, -105.288, 258.02, 2575.49, -300.668, 966.829]
  MoveL 11 to (0, 300, 221.76) mm, rotated rx 34.6 ry 1.47 rz 88.32 deg; joints [-70.837, 65.626, 6.853, -11.812, -100.438, 257.608, 2575.49, -300.668, 966.829]
  MoveL 12 to (0, 200, 222.36) mm, rotated rx 32.68 ry 1.48 rz 88.27 deg; joints [-64.457, 65.243, 2.407, -5.63, -93.694, 257.141, 2575.49, -300.668, 966.829]
  MoveL 13 to (0, 100, 223.1) mm, rotated rx 33.49 ry 1.79 rz 88.5 deg; joints [-58.749, 68.126, -6.83, -0.296, -88.008, 254.634, 2575.49, -300.668, 966.829]
  MoveL 14 to (0, 0, 224.38) mm, rotated rx 32.11 ry 1.87 rz 88.5 deg; joints [-53.551, 70.245, -16.532, 4.853, -79.401, 252.131, 2575.49, -300.668, 966.829]
  Set speed (1000.0 mm/s)
  MoveL 15 to (0, 0, 224.38) mm, rotated rx 32.11 ry 1.87 rz 88.5 deg; joints [-53.551, 70.245, -16.532, 4.853, -79.401, 252.131, 2575.49, -300.668, 966.829]
  MoveL 16 to (-53.21, -1.38, 139.72) mm, rotated rx 32.11 ry 1.87 rz 88.5 deg; joints [-50.09, 70.281, -5.521, 7.888, -90.571, 251.592, 2575.49, -300.668, 966.829]
  Set speed (1000.0 mm/s)
  MoveL 17 to (48.98, 0.77, 88.13) mm, rotated rx 15.09 ry 0.22 rz 87.5 deg; joints [-47.262, 45.262, 11.589, 13.139, -68.24, 256.627, 2575.49, -300.668, 966.829]
  MoveL 18 to (75, 0, 184.68) mm, rotated rx 15.09 ry 0.22 rz 87.5 deg; joints [-51.515, 48.761, -1.122, 9.385, -58.702, 257.474, 2575.49, -300.668, 966.829]
  MoveL 19 to (75, 0, 184.68) mm, rotated rx 15.09 ry 0.22 rz 87.5 deg; joints [-51.515, 48.761, -1.122, 9.385, -58.702, 257.474, 2575.49, -300.668, 966.829]
  Set speed (200.0 mm/s)
  MoveL 20 to (75, 100, 183.97) mm, rotated rx 14.81 ry 1.19 rz 87.75 deg; joints [-56.171, 44.891, 8.708, 4.951, -64.188, 261.236, 2575.49, -300.668, 966.829]
  MoveL 21 to (75, 200, 182.99) mm, rotated rx 14.67 ry 1.11 rz 87.73 deg; joints [-62.214, 41.805, 17.002, -1.663, -69.164, 265.152, 2575.49, -300.668, 966.829]
  MoveL 22 to (75, 300, 182.2) mm, rotated rx 14.84 ry 0.95 rz 87.69 deg; joints [-69.111, 39.859, 23.363, -8.854, -73.998, 268.206, 2575.49, -300.668, 966.829]
  MoveL 23 to (75, 400, 181.72) mm, rotated rx 15.14 ry 0.85 rz 87.67 deg; joints [-76.676, 38.911, 27.758, -16.412, -78.316, 270.529, 2575.49, -300.668, 966.829]
  MoveL 24 to (75, 500, 181.5) mm, rotated rx 15.59 ry 0.71 rz 87.63 deg; joints [-84.768, 38.925, 30.095, -24.402, -81.973, 272.402, 2575.49, -300.668, 966.829]
  MoveL 25 to (75, 600, 182.1) mm, rotated rx 15.71 ry 0.04 rz 87.44 deg; joints [-93.426, 39.497, 29.951, -33.495, -83.984, 274.919, 2575.49, -300.668, 966.829]
  MoveL 26 to (75, 700, 182.69) mm, rotated rx 18.36 ry 0.6 rz 87.62 deg; joints [-100.987, 42.892, 28.041, -39.909, -88.935, 274.72, 2575.49, -300.668, 966.829]
  MoveL 27 to (75, 800, 189.28) mm, rotated rx 49.19 ry -8.54 rz 77.42 deg; joints [-111.401, 70.498, -12.923, -60.218, -108.495, 268.047, 2575.49, -300.668, 966.829]
  MoveL 28 to (75, 900, 199.48) mm, rotated rx 34.43 ry 0.88 rz 87.91 deg; joints [-113.27, 61.136, 7.803, -49.801, -104.447, 271.342, 2575.49, -300.668, 966.829]
  MoveL 29 to (75, 1000, 185) mm, rotated rx 17 ry 0.07 rz 87.45 deg; joints [-122.024, 48.934, 10.811, -60.382, -87.552, 289.491, 2575.49, -300.668, 966.829]
  Set speed (1000.0 mm/s)
  MoveL 30 to (75, 1000, 185) mm, rotated rx 17 ry 0.07 rz 87.45 deg; joints [-122.024, 48.934, 10.811, -60.382, -87.552, 289.491, 2575.49, -300.668, 966.829]
  MoveL 31 to (45.79, 1001.19, 89.37) mm, rotated rx 17 ry 0.07 rz 87.45 deg; joints [-125.938, 46.929, 23.266, -64.051, -93.899, 281.027, 2575.49, -300.668, 966.829]
  Set speed (1000.0 mm/s)
  MoveL 32 to (131.22, 1001.22, 68.71) mm, rotated rx 10.84 ry -0.22 rz 87.42 deg; joints [-127.502, 33.7, 23.114, -67.676, -84.084, 296.685, 2575.49, -300.668, 966.829]
  MoveL 33 to (150, 1000, 166.93) mm, rotated rx 10.84 ry -0.22 rz 87.42 deg; joints [-123.243, 38.206, 10.582, -65.245, -78.512, 303.082, 2575.49, -300.668, 966.829]
  MoveL 34 to (150, 1000, 166.93) mm, rotated rx 10.84 ry -0.22 rz 87.42 deg; joints [-123.243, 38.206, 10.582, -65.245, -78.512, 303.082, 2575.49, -300.668, 966.829]
  Set speed (200.0 mm/s)
  MoveL 35 to (150, 900, 165.78) mm, rotated rx 10.61 ry 0.09 rz 87.48 deg; joints [-116.882, 33.938, 18.43, -59.03, -76.279, 297.992, 2575.49, -300.668, 966.829]
  MoveL 36 to (150, 800, 164.89) mm, rotated rx 10.45 ry 0.11 rz 87.48 deg; joints [-109.81, 30.675, 24.02, -52.243, -73.986, 293.646, 2575.49, -300.668, 966.829]
  MoveL 37 to (150, 700, 164.31) mm, rotated rx 10.08 ry 0.26 rz 87.51 deg; joints [-101.945, 28.063, 27.723, -44.556, -71.006, 289.848, 2575.49, -300.668, 966.829]
  MoveL 38 to (150, 600, 164.04) mm, rotated rx 9.89 ry 0.39 rz 87.53 deg; joints [-93.578, 26.556, 29.404, -36.164, -67.9, 285.979, 2575.49, -300.668, 966.829]
  MoveL 39 to (150, 500, 164.05) mm, rotated rx 9.84 ry 0.58 rz 87.57 deg; joints [-84.993, 26.198, 29.075, -27.229, -64.683, 281.817, 2575.49, -300.668, 966.829]
  MoveL 40 to (150, 400, 164.38) mm, rotated rx 9.61 ry 0.73 rz 87.59 deg; joints [-76.645, 26.805, 26.604, -18.368, -60.86, 277.636, 2575.49, -300.668, 966.829]
  MoveL 41 to (150, 300, 165.02) mm, rotated rx 9.43 ry 0.88 rz 87.62 deg; joints [-68.839, 28.529, 22.136, -9.632, -56.866, 272.976, 2575.49, -300.668, 966.829]
  MoveL 42 to (150, 200, 165.9) mm, rotated rx 9.44 ry 0.93 rz 87.62 deg; joints [-61.866, 31.398, 15.794, -1.341, -52.984, 267.771, 2575.49, -300.668, 966.829]
  MoveL 43 to (150, 100, 166.63) mm, rotated rx 9.53 ry 0.78 rz 87.6 deg; joints [-55.832, 35.205, 7.667, 6.348, -48.92, 262.124, 2575.49, -300.668, 966.829]
  MoveL 44 to (150, 0, 166.55) mm, rotated rx 9.95 ry 0.36 rz 87.53 deg; joints [-50.719, 39.991, -2.111, 13.391, -44.944, 255.947, 2575.49, -300.668, 966.829]
  Set speed (1000.0 mm/s)
  MoveL 45 to (150, 0, 166.55) mm, rotated rx 9.95 ry 0.36 rz 87.53 deg; joints [-50.719, 39.991, -2.111, 13.391, -44.944, 255.947, 2575.49, -300.668, 966.829]
  MoveL 46 to (132.71, 0.12, 68.05) mm, rotated rx 9.95 ry 0.36 rz 87.53 deg; joints [-46.21, 34.77, 10.454, 17.523, -52.918, 254.226, 2575.49, -300.668, 966.829]
  Set speed (1000.0 mm/s)
  MoveL 47 to (217.88, 1.74, 58.04) mm, rotated rx 4.12 ry -0.82 rz 87.44 deg; joints [-46.796, 26.316, 4.174, 22.706, -33.753, 250.007, 2575.49, -300.668, 966.829]
  MoveL 48 to (225, 0, 157.77) mm, rotated rx 4.12 ry -0.82 rz 87.44 deg; joints [-51.251, 33.338, -8.257, 17.496, -27.319, 253.636, 2575.49, -300.668, 966.829]
  MoveL 49 to (225, 0, 157.77) mm, rotated rx 4.12 ry -0.82 rz 87.44 deg; joints [-51.251, 33.338, -8.257, 17.496, -27.319, 253.636, 2575.49, -300.668, 966.829]
  Set speed (200.0 mm/s)
  MoveL 50 to (225, 100, 158.69) mm, rotated rx 4.01 ry -0.16 rz 87.49 deg; joints [-56.364, 28.112, 1.373, 6.828, -30.708, 263.57, 2575.49, -300.668, 966.829]
  MoveL 51 to (225, 200, 158.45) mm, rotated rx 3.23 ry 0.33 rz 87.52 deg; joints [-62.286, 23.428, 8.777, -3.628, -32.63, 272.978, 2575.49, -300.668, 966.829]
  MoveL 52 to (225, 300, 157.75) mm, rotated rx 3.35 ry 0.61 rz 87.54 deg; joints [-69.113, 19.975, 15.018, -14.433, -36.344, 281.636, 2575.49, -300.668, 966.829]
  MoveL 53 to (225, 400, 157.18) mm, rotated rx 3.55 ry 0.49 rz 87.53 deg; joints [-76.99, 17.692, 19.433, -25.79, -40.748, 290.05, 2575.49, -300.668, 966.829]
  MoveL 54 to (225, 500, 156.9) mm, rotated rx 3.54 ry 0.3 rz 87.52 deg; joints [-85.455, 16.603, 21.74, -36.696, -45.337, 297.703, 2575.49, -300.668, 966.829]
  MoveL 55 to (225, 600, 156.89) mm, rotated rx 3.67 ry 0.16 rz 87.51 deg; joints [-94.073, 16.916, 22.192, -46.262, -50.533, 303.788, 2575.49, -300.668, 966.829]
  MoveL 56 to (225, 700, 157.17) mm, rotated rx 3.64 ry -0.01 rz 87.5 deg; joints [-102.526, 18.492, 20.531, -54.974, -55.638, 309.21, 2575.49, -300.668, 966.829]
  MoveL 57 to (225, 800, 157.75) mm, rotated rx 3.62 ry -0.18 rz 87.49 deg; joints [-110.436, 21.291, 16.897, -62.522, -60.59, 313.924, 2575.49, -300.668, 966.829]
  MoveL 58 to (225, 900, 158.59) mm, rotated rx 3.75 ry -0.5 rz 87.47 deg; joints [-117.643, 25.324, 11.226, -69.016, -65.45, 318.24, 2575.49, -300.668, 966.829]
  MoveL 59 to (225, 1000, 159.66) mm, rotated rx 3.77 ry -0.44 rz 87.47 deg; joints [-123.843, 30.006, 3.902, -74.249, -69.389, 322.651, 2575.49, -300.668, 966.829]
  Set speed (1000.0 mm/s)
  MoveL 60 to (225, 1000, 159.66) mm, rotated rx 3.77 ry -0.44 rz 87.47 deg; joints [-123.843, 30.006, 3.902, -74.249, -69.389, 322.651, 2575.49, -300.668, 966.829]
  MoveL 61 to (218.47, 1001.06, 59.88) mm, rotated rx 3.77 ry -0.44 rz 87.47 deg; joints [-128.254, 23.194, 15.755, -75.572, -74.131, 318.504, 2575.49, -300.668, 966.829]
  Set speed (1000.0 mm/s)
  MoveL 62 to (300.78, 1001, 58.22) mm, rotated rx -0.42 ry -0.59 rz 87.53 deg; joints [-128.379, 18.573, 5.193, -83.874, -69.705, 337.428, 2575.49, -300.668, 966.829]
  MoveL 63 to (300, 1000, 158.21) mm, rotated rx -0.42 ry -0.59 rz 87.53 deg; joints [-123.978, 26.422, -6.075, -83.441, -65.272, 340.615, 2575.49, -300.668, 966.829]
  MoveL 64 to (300, 1000, 158.21) mm, rotated rx -0.42 ry -0.59 rz 87.53 deg; joints [-123.978, 26.422, -6.075, -83.441, -65.272, 340.615, 2575.49, -300.668, 966.829]
  Set speed (200.0 mm/s)
  MoveL 65 to (300, 900, 157.2) mm, rotated rx -0.44 ry -0.43 rz 87.53 deg; joints [-117.734, 21.144, 1.519, -79.458, -59.714, 337.05, 2575.49, -300.668, 966.829]
  MoveL 66 to (300, 800, 156.45) mm, rotated rx -0.59 ry -0.48 rz 87.53 deg; joints [-110.757, 17.059, 6.67, -75.266, -53.678, 334.296, 2575.49, -300.668, 966.829]
  MoveL 67 to (300, 700, 155.94) mm, rotated rx -0.69 ry -0.34 rz 87.53 deg; joints [-102.947, 14.033, 10.076, -70.036, -46.808, 331.121, 2575.49, -300.668, 966.829]
  MoveL 68 to (300, 600, 155.62) mm, rotated rx -0.64 ry -0.19 rz 87.53 deg; joints [-94.596, 12.369, 11.692, -63.29, -39.686, 326.634, 2575.49, -300.668, 966.829]
  MoveL 69 to (300, 500, 155.56) mm, rotated rx -0.7 ry -0.06 rz 87.53 deg; joints [-86.037, 12.123, 11.29, -55.019, -32.482, 320.74, 2575.49, -300.668, 966.829]
  MoveL 70 to (300, 400, 155.72) mm, rotated rx -0.76 ry 0.06 rz 87.52 deg; joints [-77.658, 13.334, 8.989, -44.15, -25.758, 312.106, 2575.49, -300.668, 966.829]
  MoveL 71 to (300, 300, 156.14) mm, rotated rx -0.69 ry 0.29 rz 87.52 deg; joints [-69.703, 15.943, 4.897, -28.595, -20.057, 298.484, 2575.49, -300.668, 966.829]
  MoveL 72 to (300, 200, 156.6) mm, rotated rx 0.08 ry 0.05 rz 87.52 deg; joints [-62.801, 19.92, -0.487, -9.383, -17.296, 280.349, 2575.49, -300.668, 966.829]
  MoveL 73 to (300, 100, 156.28) mm, rotated rx 0.08 ry -0.57 rz 87.52 deg; joints [-56.912, 24.724, -8.418, 10.218, -14.184, 261.712, 2575.49, -300.668, 966.829]
  MoveL 74 to (300, 0, 154.7) mm, rotated rx 0.72 ry -1.11 rz 87.5 deg; joints [-51.648, 30.572, -17.827, 33.669, -13.102, 238.455, 2575.49, -300.668, 966.829]
  Set speed (1000.0 mm/s)
  MoveL 75 to (300, 0, 154.7) mm, rotated rx 0.72 ry -1.11 rz 87.5 deg; joints [-51.648, 30.572, -17.827, 33.669, -13.102, 238.455, 2575.49, -300.668, 966.829]
  MoveL 76 to (298.82, 2, 54.73) mm, rotated rx 0.72 ry -1.11 rz 87.5 deg; joints [-47.249, 22.565, -5.438, 37.879, -19.143, 235.259, 2575.49, -300.668, 966.829]
  Set speed (1000.0 mm/s)
  MoveL 77 to (377.68, 2.79, 55.06) mm, rotated rx -1.47 ry -1.66 rz 87.57 deg; joints [-48.108, 21.555, -17.026, 85.224, -10.172, 187.886, 2575.49, -300.668, 966.829]
  MoveL 78 to (375, 0, 154.99) mm, rotated rx -1.47 ry -1.66 rz 87.57 deg; joints [-52.369, 30.453, -30.168, 119.554, -6.767, 153.034, 2575.49, -300.668, 966.829]
  MoveL 79 to (375, 0, 154.99) mm, rotated rx -1.47 ry -1.66 rz 87.57 deg; joints [-52.369, 30.453, -30.168, 119.554, -6.767, 153.034, 2575.49, -300.668, 966.829]
  Set speed (200.0 mm/s)
  MoveL 80 to (375, 100, 157.33) mm, rotated rx -1.72 ry -0.53 rz 107.55 deg; joints [-56.618, 25.011, -10.257, 11.369, -21.322, 278.684, 2575.49, -300.668, 966.829]
  MoveL 81 to (375, 200, 158.25) mm, rotated rx -2.25 ry -0.49 rz 87.55 deg; joints [-63.645, 19.043, -12.028, -57.753, -5, 330.046, 2575.49, -300.668, 966.829]
  MoveL 82 to (375, 300, 158.07) mm, rotated rx -2.21 ry 0.1 rz 87.53 deg; joints [-70.28, 14.985, -5.746, -64.97, -11.324, 336.4, 2575.49, -300.668, 966.829]
  MoveL 83 to (375, 400, 157.85) mm, rotated rx -2.55 ry -0.08 rz 87.54 deg; joints [-78.166, 12.265, -1.942, -73.941, -19.069, 344.37, 2575.49, -300.668, 966.829]
  MoveL 84 to (375, 500, 157.83) mm, rotated rx -2.47 ry -0.14 rz 87.54 deg; joints [-86.424, 10.961, 0.429, -77.607, -27.266, 346.638, 2575.49, -300.668, 966.829]
  MoveL 85 to (375, 600, 157.94) mm, rotated rx -2.9 ry -0.27 rz 87.55 deg; joints [-94.885, 11.163, 0.297, -82.3, -35.505, 350.14, 2575.49, -300.668, 966.829]
  MoveL 86 to (375, 700, 158.26) mm, rotated rx -2.95 ry -0.42 rz 87.56 deg; joints [-103.132, 12.863, -1.316, -85.028, -43.688, 351.509, 2575.49, -300.668, 966.829]
  MoveL 87 to (375, 800, 158.82) mm, rotated rx -3 ry -0.55 rz 87.57 deg; joints [-110.832, 15.957, -4.888, -87.513, -51.316, 352.905, 2575.49, -300.668, 966.829]
  MoveL 88 to (375, 900, 159.55) mm, rotated rx -2.84 ry -0.6 rz 87.57 deg; joints [-117.769, 20.278, -10.219, -89.461, -58.174, 354.179, 2575.49, -300.668, 966.829]
  MoveL 89 to (375, 1000, 160.39) mm, rotated rx -2.82 ry -0.6 rz 87.57 deg; joints [-123.887, 25.771, -17.978, -91.612, -64.238, 356.682, 2575.49, -300.668, 966.829]
  Set speed (1000.0 mm/s)
  MoveL 90 to (375, 1000, 160.39) mm, rotated rx -2.82 ry -0.6 rz 87.57 deg; joints [-123.887, 25.771, -17.978, -91.612, -64.238, 356.682, 2575.49, -300.668, 966.829]
  MoveL 91 to (379.97, 1000.83, 60.52) mm, rotated rx -2.82 ry -0.6 rz 87.57 deg; joints [-128.216, 17.356, -6.724, -91.018, -68.446, 353.478, 2575.49, -300.668, 966.829]
  Set speed (1000.0 mm/s)
  MoveL 92 to (440.72, 900.9, 61.47) mm, rotated rx 5.34 ry -0.28 rz 87.47 deg; joints [-121.633, 11.757, 1.394, -80.715, -63.31, 342.925, 2575.49, -300.668, 966.829]
  MoveL 93 to (450, 900, 161.03) mm, rotated rx 5.34 ry -0.28 rz 87.47 deg; joints [-117.735, 20.445, -11.137, -81.729, -58.942, 346.594, 2575.49, -300.668, 966.829]
  MoveL 94 to (450, 900, 161.03) mm, rotated rx 5.34 ry -0.28 rz 87.47 deg; joints [-117.735, 20.445, -11.137, -81.729, -58.942, 346.594, 2575.49, -300.668, 966.829]
  Set speed (200.0 mm/s)
  MoveL 95 to (450, 800, 160.5) mm, rotated rx 5.21 ry -0.05 rz 87.49 deg; joints [-110.719, 15.993, -5.562, -79.024, -52.059, 343.947, 2575.49, -300.668, 966.829]
  MoveL 96 to (450, 700, 160.24) mm, rotated rx 4.96 ry 0.1 rz 87.5 deg; joints [-103.01, 12.906, -2.334, -76.267, -44.477, 341.866, 2575.49, -300.668, 966.829]
  MoveL 97 to (450, 600, 160.2) mm, rotated rx 4.56 ry 0.21 rz 87.51 deg; joints [-94.8, 11.236, -1.26, -73.435, -36.306, 340.032, 2575.49, -300.668, 966.829]
  MoveL 98 to (450, 500, 160.37) mm, rotated rx 4.48 ry 0.35 rz 87.52 deg; joints [-86.36, 11.076, -1.759, -68.74, -28.059, 336.202, 2575.49, -300.668, 966.829]
  MoveL 99 to (450, 400, 160.59) mm, rotated rx -0.82 ry 0.05 rz 87.52 deg; joints [-78.425, 12.602, -10.427, -93.358, -18.429, 364.448, 2575.49, -300.668, 966.829]
  MoveL 100 to (450, 300, 160.76) mm, rotated rx -0.75 ry 0.08 rz 87.52 deg; joints [-70.692, 15.45, -14.739, -102.619, -10.914, 374.181, 2575.49, -300.668, 966.829]
  MoveL 101 to (450, 200, 160.9) mm, rotated rx -0.33 ry 0.18 rz 107.52 deg; joints [-62.593, 19.724, -10.529, -2.747, -16.272, 291.889, 2575.49, -300.668, 966.829]
  MoveL 102 to (450, 100, 160.1) mm, rotated rx -2.38 ry -0.56 rz 107.57 deg; joints [-57.222, 24.711, -20.554, 18.628, -10.342, 271.393, 2575.49, -300.668, 966.829]
  MoveL 103 to (450, 0, 157.34) mm, rotated rx -2.09 ry -2.03 rz 87.61 deg; joints [-53.037, 32.949, -45.422, 163.573, -17.277, 108.816, 2575.49, -300.668, 966.829]
  Set speed (1000.0 mm/s)
  MoveL 104 to (450, 0, 157.34) mm, rotated rx -2.09 ry -2.03 rz 87.61 deg; joints [-53.037, 32.949, -45.422, 163.573, -17.277, 108.816, 2575.49, -300.668, 966.829]
  MoveL 105 to (453.79, 3.39, 57.47) mm, rotated rx -2.09 ry -2.03 rz 87.61 deg; joints [-48.895, 22.769, -29.81, 141.003, -14.312, 131.511, 2575.49, -300.668, 966.829]
  Set speed (1000.0 mm/s)
  MoveL 106 to (509.65, -0.21, 55.44) mm, rotated rx 8.81 ry 0.5 rz 87.55 deg; joints [-47.244, 23.046, -25.215, 76.548, -13.462, 189.728, 2575.49, -300.668, 966.829]
  MoveL 107 to (525, 0, 154.26) mm, rotated rx 8.81 ry 0.5 rz 87.55 deg; joints [-51.722, 32.801, -42.664, 117.795, -9.763, 148.192, 2575.49, -300.668, 966.829]
  MoveL 108 to (525, 0, 154.26) mm, rotated rx 8.81 ry 0.5 rz 87.55 deg; joints [-51.722, 32.801, -42.664, 117.795, -9.763, 148.192, 2575.49, -300.668, 966.829]
  Set speed (200.0 mm/s)
  MoveL 109 to (525, 100, 153.45) mm, rotated rx 10.33 ry 0.99 rz 87.65 deg; joints [-56.932, 25.038, -27.321, 42.012, -5.764, 224.113, 2575.49, -300.668, 966.829]
  MoveL 110 to (525, 200, 152.5) mm, rotated rx 10.55 ry 1.07 rz 87.66 deg; joints [-63.114, 19.275, -17.751, -15.039, -8.572, 281.466, 2575.49, -300.668, 966.829]
  MoveL 111 to (525, 300, 151.54) mm, rotated rx 9.35 ry 0.76 rz 87.59 deg; joints [-70.339, 14.873, -12.407, -49.938, -12.679, 317.099, 2575.49, -300.668, 966.829]
  MoveL 112 to (525, 400, 150.88) mm, rotated rx 8.9 ry 0.66 rz 87.58 deg; joints [-78.153, 11.939, -8.476, -63.621, -19.653, 331.006, 2575.49, -300.668, 966.829]
  MoveL 113 to (525, 500, 150.43) mm, rotated rx 8.39 ry 0.49 rz 87.55 deg; joints [-86.519, 10.508, -6.658, -71.794, -27.517, 339.365, 2575.49, -300.668, 966.829]
  MoveL 114 to (525, 600, 150.24) mm, rotated rx 7.97 ry 0.34 rz 87.52 deg; joints [-95.026, 10.628, -6.689, -76.729, -35.747, 344.434, 2575.49, -300.668, 966.829]
  MoveL 115 to (525, 700, 150.34) mm, rotated rx 7.96 ry 0.25 rz 87.51 deg; joints [-103.27, 12.276, -8.186, -79.237, -43.904, 346.92, 2575.49, -300.668, 966.829]
  MoveL 116 to (525, 800, 150.74) mm, rotated rx 7.62 ry 0.05 rz 87.49 deg; joints [-111.05, 15.453, -12.171, -82.05, -51.581, 350.162, 2575.49, -300.668, 966.829]
  MoveL 117 to (525, 900, 151.36) mm, rotated rx 7.45 ry -0.12 rz 87.46 deg; joints [-118.056, 20.016, -18.197, -84.174, -58.504, 353.16, 2575.49, -300.668, 966.829]
  Set speed (1000.0 mm/s)
  MoveL 118 to (525, 900, 151.36) mm, rotated rx 7.45 ry -0.12 rz 87.46 deg; joints [-118.056, 20.016, -18.197, -84.174, -58.504, 353.16, 2575.49, -300.668, 966.829]
  MoveL 119 to (512.06, 900.79, 52.2) mm, rotated rx 7.45 ry -0.12 rz 87.46 deg; joints [-121.985, 11.006, -4.868, -82.299, -62.909, 348.775, 2575.49, -300.668, 966.829]

--- program DoorFR (robot ABB IRB 1300-10/1.15) ---
  Smooth(1)
  Set speed (1000.0 mm/s)
  Set Ref.: DoorFR
  Set Tool: Generic Paint Sprayer
  Show Generic Paint Sprayer
  MoveJ 1 to (-16.42, 1.32, 177.76) mm, rotated rx 9.47 ry -0.34 rz 87.41 deg; joints [-50.928, 50.766, 2.133, 9.955, -59.087, 260.693, 2575.49, -300.668, 966.829]
  MoveL 2 to (-16.42, 1.32, 177.76) mm, rotated rx 9.47 ry -0.34 rz 87.41 deg; joints [-50.928, 50.766, 2.133, 9.955, -59.087, 260.693, 2575.49, -300.668, 966.829]
  MoveL 3 to (0, 0, 276.4) mm, rotated rx 9.47 ry -0.34 rz 87.41 deg; joints [-54.628, 55.899, -12.659, 6.412, -49.179, 262.02, 2575.49, -300.668, 966.829]
  MoveL 4 to (0, 0, 276.4) mm, rotated rx 9.47 ry -0.34 rz 87.41 deg; joints [-54.628, 55.899, -12.659, 6.412, -49.179, 262.02, 2575.49, -300.668, 966.829]
  Set speed (20.0 mm/s)
  MoveL 5 to (0, 100, 332.15) mm, rotated rx 43.66 ry 50.93 rz -91.45 deg; joints [-87.183, 40.143, -38.431, 193.477, -38.824, 229.231, 3075.49, -300.668, 966.829]
  Set speed (1000.0 mm/s)
  MoveL 6 to (0, 100, 332.15) mm, rotated rx 17.45 ry 61.45 rz -122.62 deg; joints [-90.156, 36.935, -25.016, 221.544, -26.283, 183.935, 3075.49, -300.668, 966.829]
  MoveL 7 to (70.43, 154.41, 286.56) mm, rotated rx 17.45 ry 61.45 rz -122.62 deg; joints [-93.916, 31.766, -25.341, 219.616, -32.87, 185.46, 3075.49, -300.668, 966.829]

